RoboDK station: Componentes_Grupo4.rdk

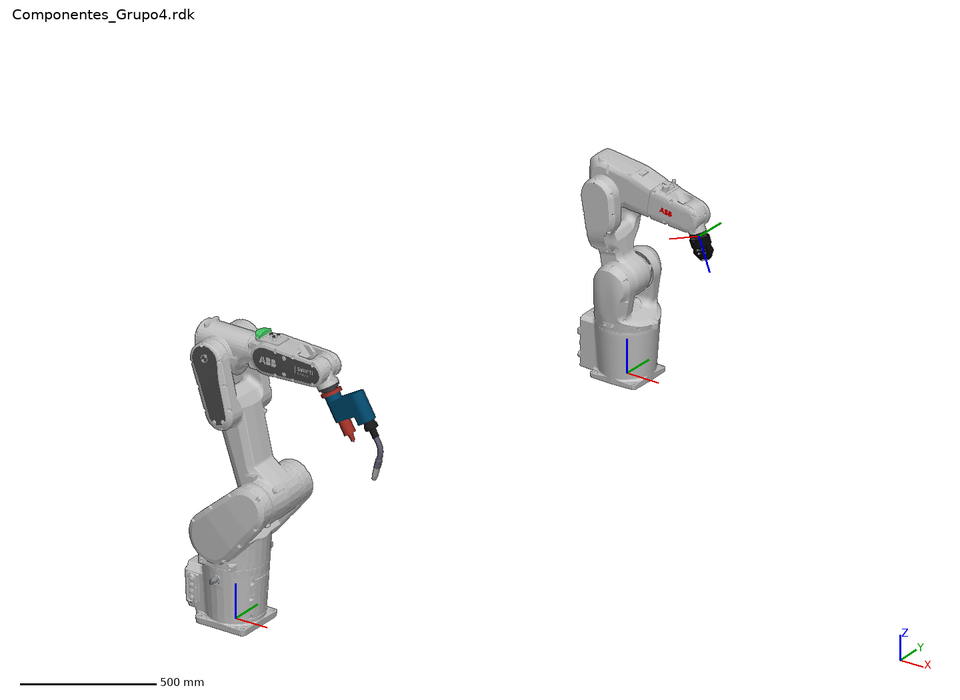
[picture v0: the station drawn from its stored meshes, robots at their saved joint values, targets as dots, program paths as lines]
Station Componentes_Grupo4 (saved by RoboDK 6.1.1). Poses are relative to the parent item; angles as X-Y-Z fixed-axis rotations.
  - frame ABB CRB 1300-10/1.15 Base at (0, 0, 0) mm
    - robot ABB CRB 1300-10/1.15: 6 axes
        modified DH rows (alpha deg, a mm, theta deg, d mm): 0, 0, 0, 544; -90, 150, -90, 0; 0, 575, 0, 0; -90, 40, 0, 425; 90, 0, 0, 0; -90, 0, 180, 90
        joint limits [-180, -95, -210, -230, -130, -242] to [180, 155, 65, 230, 130, 242]; home [0, 0, 0, 0, 0, 0]; saved at [0, -20, 20, 0, 60, 0]
      - tool Generic Welding Gun (Over-arm), TCP at (-4, 0, 371.3) mm, rotated rx 0 ry 45 rz 0 deg, size 169.7 x 60 x 367 mm
      - tool Antorcha_TIG, TCP at (0, 0, 207) mm, size 80 x 80 x 207 mm, geometry from antorcha_tig.stl
  - frame ABB IRB 1200-7/0.7 Base at (0, 2500, 0) mm
    - robot ABB IRB 1200-7/0.7: 6 axes, payload 7 kg, reach 703 mm, repeatability 0.02 mm, weight 54 kg
        modified DH rows (alpha deg, a mm, theta deg, d mm): 0, 0, 0, 399; -90, 0, -90, 0; 0, 350, 0, 0; -90, 42, 0, 351; 90, 0, 0, 0; -90, 0, 180, 82
        joint limits [-170, -100, -200, -270, -130, -360] to [170, 135, 70, 270, 130, 360]; home [0, 0, 0, 0, 0, 0]; saved at [0, -10, 20, 0, 60, 0]
      - frame RobotiQ 2F-85 Gripper (Mechanism) Base at (0, 0, 0) mm
        - robot RobotiQ 2F-85 Gripper (Mechanism) (model RobotiQ 2F85): 1 axes, payload 5 kg
            joint limits [0] to [85]; home [85]; saved at [85]
  - object paquete_estator at (0, 5000, 0) mm, size 105 x 105 x 55 mm, geometry from paquete_estator.stl
  - object pallet_4_posiciones at (0, 7000, 0) mm, size 400 x 400 x 20 mm, geometry from pallet_4_posiciones.stl
  - frame ConveyorA Base at (6000, 0, 0) mm
    - robot ConveyorA: 1 axes
        modified DH rows (alpha deg, a mm, theta deg, d mm): 0, 0, 0, 0 linear
        base shift (0, 0, 0) mm, rotated rx 0 ry 90 rz 0 deg
        joint limits [-900000] to [900000]; home [0]; saved at [0]
  - object Laser-Sensor at (6000, 4000, 0) mm, size 683.3 x 45.2 x 12.5 mm, geometry from Laser-Sensor.stl
  - object Table-1400x800x800mm at (6000, 8000, 0) mm, size 1420 x 820 x 800 mm, geometry from Table-1400x800x800mm.stl
  - object estacion_servicio_antorcha at (0, -3000, 0) mm, size 250 x 250 x 1000 mm, geometry from estacion_servicio_antorcha.stl
